Fanuc KAREL source: ka00001.KL

PROGRAM KA00001
%STACKSIZE=65535
%PRIORITY=65535
%NOLOCKGROUP
VAR
SRC : INTEGER
DST : INTEGER
BEGIN
SRC=2
DST=SRC
END KA00001
